// TIA Portal V19 export
DATA_BLOCK "Tacho2_EM01"   // DB2
VERSION : 1.0
// stored: InstanceOfName EM01_Calentamiento, InstanceOfType FB
"EM01_Calentamiento"
   // VAR_INPUT
   //    In : "EM01_Input";
   //    TempPV : Real;
   //    TempValid : Bool;
   //    ConcPV : Real;
   //    ConcValid : Bool;
   // END_VAR
   // VAR_OUTPUT
   //    Out : "EM01_Output";
   //    CM_Out : Bool;
   //    CM_Pid_MV : Real;
   // END_VAR
   // VAR
   //    State : Int;
   //    FaultLatched : Bool;
   //    FaultCode : Int;
   //    ActiveMode : Int;
   //    ElapsedPrev : Time;
   //    TimerConc { S7_SetPoint := 'True'} : TON_TIME;
   //    TimerTemp { S7_SetPoint := 'True'} : TON_TIME;
   //    TimerTime { S7_SetPoint := 'True'} : TON_TIME;
   //    TimerFault { S7_SetPoint := 'True'} : TON_TIME;
   //    TimerOpen { S7_SetPoint := 'True'} : TON_TIME;
   //    TimerClose { S7_SetPoint := 'True'} : TON_TIME;
   //    TrigStart { S7_SetPoint := 'True'} : R_TRIG;
   //    TrigStop { S7_SetPoint := 'True'} : R_TRIG;
   //    TrigHold { S7_SetPoint := 'True'} : R_TRIG;
   //    TrigAbort { S7_SetPoint := 'True'} : R_TRIG;
   //    TrigReset { S7_SetPoint := 'True'} : R_TRIG;
   //    CM_Vlv_Cal { S7_SetPoint := 'True'} : "VlvL";   // Valv
   //    CM_Pid_CalandriaVapor { S7_SetPoint := 'True'} : "PidL";   // PID
   // END_VAR
BEGIN
   CM_Vlv_Cal.DataHMI.identName := 'V1';
   CM_Vlv_Cal.DataHMI.comment := 'Calentamiento';
   CM_Pid_CalandriaVapor.PV_unit := 1426;
   CM_Pid_CalandriaVapor.DataHMI.identName := 'DIC';
   CM_Pid_CalandriaVapor.DataHMI.comment := 'Concentracion';
END_DATA_BLOCK
